ABB RAPID module: PickIn1.mod

%%%
  VERSION:1
  LANGUAGE:ENGLISH
%%%
MODULE MOD_PickIn1

    ! -------------------------------
    ! Define customized variables here
    ! ...

	! Tool variables:
	PERS tooldata SuctionCup := [TRUE,[[-94.709,0.000,259.352],[0.00000000,0.00000000,0.00000000,1.00000000]],[1,[0,0,20],[1,0,0,0],0,0,0.005]];

	! Reference variables:
	PERS wobjdata In := [FALSE, TRUE, "", [[0,0,0],[1,0,0,0]],[[290.000,450.000,10.000],[1.00000000,0.00000000,0.00000000,0.00000000]]];

	PROC Main()
		ConfJ \On;
		ConfL \Off;
		! Program generated by VerticalBot Studio for ABB IRB 1200-5/0.9 on 25/10/2026 12:00:00
		! Using nominal kinematics.
		MoveAbsJ [[70.152800,32.938500,23.515600,0.000000,33.545900,70.152800],[9E+09,9E+09,9E+09,9E+09,9E+09,9E+09]],v500,z1,SuctionCup \WObj:=In;
		MoveL [[-16.111,46.392,45.000],[0.00000000,1.00000000,0.00000000,-0.00000000],[0,2,-2,1],[9E+09,9E+09,9E+09,9E+09,9E+09,9E+09]],v500,z1,SuctionCup \WObj:=In;
		! Attach to Suction Cup
		WaitTime 0.500;
		MoveL [[-16.087,46.472,70.960],[0.00000000,1.00000000,0.00000000,-0.00000000],[0,0,0,0],[9E+09,9E+09,9E+09,9E+09,9E+09,9E+09]],v500,z1,SuctionCup \WObj:=In;
	ENDPROC

ENDMODULE
